Fanuc KAREL source: KT00706.KL

PROGRAM KT00706
%NOLOCKGROUP
VAR
  I1: INTEGER
  I2: INTEGER
  OUT: BOOLEAN
BEGIN
  I1 = 2
  I2 = 3
  I1 = 2
  I2 = 3
  OUT = UNINIT(I1)
END KT00706
